SUBAPPLICATION SubApp_PC_B (* Geraet B: Flip-Flop (opcua.adoc): SUBSCRIBE Flip -> E_SWITCH/E_SR -> PUBLISH Flop; Input_I1 schreibt Flip, Output_Q1 zeigt Flop (= NICHT I1) *)
  (* Standard: 61499-2; Description: Copyright (c) 2026 Meisterschulen am Ostbahnhof This program and the accompanying materials are made available under the terms of the Eclipse Public License 2.0 which is available at https://www.eclipse.org/legal/epl-2.0/ SPDX-License-Identifier: EPL-2.0 *)
  (* Version 1.0, 2026-10-18, Franz Höpfinger, Meisterschulen am Ostbahnhof, opcua.adoc-Beispiel auf zwei Geraeten *)
  PACKAGE subapp::Training_13_OPC_UA_RES;
  IMPORT VV::const::OPC_UA::myOpcUaAddresses::T13_FLIP_READ;
  IMPORT VV::const::OPC_UA::myOpcUaAddresses::T13_FLOP_WRITE;
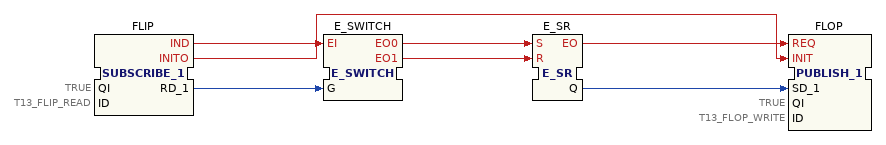
  FBS
    FLIP : iec61499::net::SUBSCRIBE_1(QI := TRUE, ID := T13_FLIP_READ);
    E_SWITCH : iec61499::events::E_SWITCH;
    E_SR : iec61499::events::E_SR;
    FLOP : iec61499::net::PUBLISH_1(QI := TRUE, ID := T13_FLOP_WRITE);
  END_FBS
  EVENT_CONNECTIONS
    FLIP.IND TO E_SWITCH.EI;
    E_SWITCH.EO0 TO E_SR.S;
    E_SWITCH.EO1 TO E_SR.R;
    E_SR.EO TO FLOP.REQ;
    FLIP.INITO TO FLOP.INIT;
  END_CONNECTIONS
  DATA_CONNECTIONS
    FLIP.RD_1 TO E_SWITCH.G;
    E_SR.Q TO FLOP.SD_1;
  END_CONNECTIONS
END_SUBAPPLICATION
